// CFC twin of T_SafeTon_Tests: the same tests drawn as CFC diagrams, the way a TwinSAFE project is authored.
    FUNCTION_BLOCK T_SafeTon_Tests_CFC EXTENDS T_SafeCfcTestSuite
    VAR
    // Test_OutputDelayedOn
    group_1 : T_SafeGroup;
    fb_1 : T_SafeTon(group := group_1) := (Parameters := (DelayTime := T#100MS));
    trigStart_1 : R_TRIG;
    t1_1 : TON;
    trig1_1 : R_TRIG;
END_VAR

Test_OutputDelayedOn();

METHOD PRIVATE Test_OutputDelayedOn
// note: this text did not pass the execution check against the stored diagram
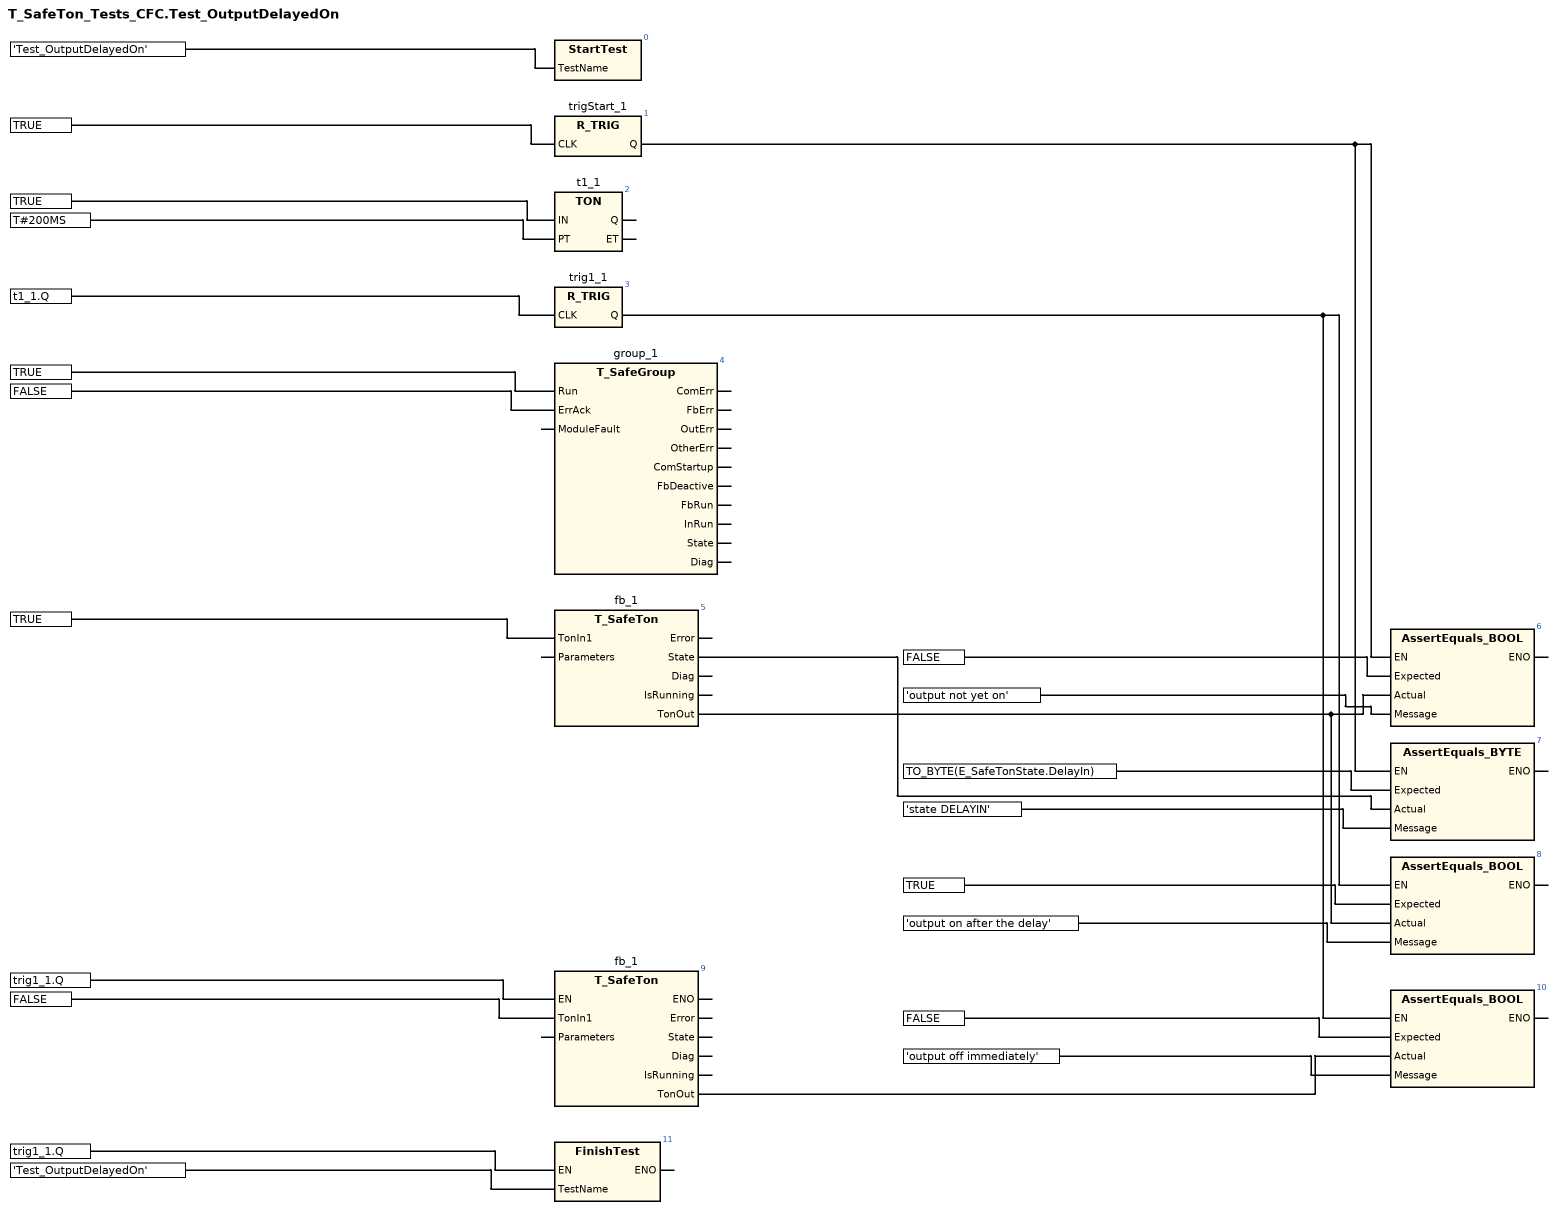
StartTest(TestName := 'Test_OutputDelayedOn');
trigStart_1(CLK := TRUE); // R_TRIG
t1_1(IN := TRUE, PT := T#200MS); // TON
trig1_1(CLK := t1_1.Q); // R_TRIG
group_1(Run := TRUE, ErrAck := FALSE); // T_SafeGroup
fb_1(TonIn1 := TRUE); // T_SafeTon
IF trigStart_1.Q THEN AssertEquals_BOOL(Expected := FALSE, Actual := fb_1.TonOut, Message := 'output not yet on'); END_IF
IF trigStart_1.Q THEN AssertEquals_BYTE(Expected := TO_BYTE(E_SafeTonState.DelayIn), Actual := fb_1.State, Message := 'state DELAYIN'); END_IF
IF trig1_1.Q THEN AssertEquals_BOOL(Expected := TRUE, Actual := fb_1.TonOut, Message := 'output on after the delay'); END_IF
IF trig1_1.Q THEN
    fb_1(TonIn1 := FALSE); // T_SafeTon
END_IF
IF trig1_1.Q THEN AssertEquals_BOOL(Expected := FALSE, Actual := fb_1.TonOut, Message := 'output off immediately'); END_IF
IF trig1_1.Q THEN FinishTest(TestName := 'Test_OutputDelayedOn'); END_IF
END_METHOD

END_FUNCTION_BLOCK

(* stored: Version 1.1.0.1, ProductVersion 3.1.4026.22
   POU T_SafeTon_Tests_CFC: Id {fb9daef6-62e7-5ece-a171-f1a002b5b4d0}, SpecialFunc None
   Method Test_OutputDelayedOn: Id {8acc0fc5-5576-5f53-a728-9d5750a35922} *)
